Staubli VAL3: getToolID.pgx

public program getToolID(string x_sKey, num& x_nToolID)
begin
   x_nToolID=trajTemp:tTrajItem[x_sKey].nToolIndex
end
